{attribute 'qualified_only'}
{attribute 'strict'}
{attribute 'to_string'}
TYPE E_Word :
(
	eOptionA := 0,
	eOptionB,
	eOptionC
) WORD;
END_TYPE

(* stored: Version 1.1.0.1, ProductVersion 3.1.4026.19
   DUT E_Word: Id {56b9148a-9331-4bb8-9b0c-9450f9ddbb2f} *)
